{attribute 'no_assign'}
FUNCTION_BLOCK FB_LN_WTURBINE_LD0_LPHD1 EXTENDS FB_AcsiCommonLogicalNodeClass
VAR_INPUT
	PhyNam: FB_DO_WTURBINE_LD0_LPHD1_PhyNam := (sClass:='WDPL', bLinkResult:=THIS^.AddDataToContainer(ipData:=PhyNam));
	PhyHealth: FB_DO_WTURBINE_LD0_LPHD1_PhyHealth := (sClass:='ENS', bLinkResult:=THIS^.AddDataToContainer(ipData:=PhyHealth));
	Proxy: FB_DO_WTURBINE_LD0_LPHD1_Proxy := (sClass:='SPS', bLinkResult:=THIS^.AddDataToContainer(ipData:=Proxy));
END_VAR
VAR
END_VAR

END_FUNCTION_BLOCK

(* stored: Version 1.1.0.1
   POU FB_LN_WTURBINE_LD0_LPHD1: Id {4f8ff99b-2dda-462b-8dba-e3f017ceb577}, SpecialFunc None *)
